(* IEC 61131-3 sources: plc-st-coding-agent/agent_dev/tests/samples, 4 files *)

(* ---- _bad_missing_clip.st ---- *)
FUNCTION_BLOCK FB
VAR_INPUT
    enable : BOOL;
    values : ARRAY[1..8] OF INT;
    count : INT;
    avgEnable : BOOL;
END_VAR
VAR_OUTPUT
    avgOut : REAL;
END_VAR
VAR
    i : INT;
    sum : DINT;
END_VAR
IF enable AND avgEnable AND count > 0 THEN
    sum := 0;
    FOR i := 1 TO count DO
        sum := sum + values[i];
    END_FOR
    avgOut := DINT_TO_REAL(sum) / INT_TO_REAL(count);
END_IF
END_FUNCTION_BLOCK

(* ---- bad_counter.st ---- *)
FUNCTION_BLOCK Bad
VAR_INPUT
    Start : BOOL;
END_VAR
VAR_OUTPUT
    Count : INT;
END_VAR
VAR
    Edge : BOOL;
END_VAR

IF Start THEN
    Count := Count + 1;
    Start := FALSE;
END_IF
IF Count > 100 THEN
    Edge := TRUE
END_IF;
IF Edge THEN
    Count := lalala + 1;
END_IF;
END_FUNCTION_BLOCK

(* ---- ok_counter.st ---- *)
FUNCTION_BLOCK Counter
VAR_INPUT
    Start : BOOL;
    Reset : BOOL;
END_VAR
VAR_OUTPUT
    Count : INT;
    Running : BOOL;
END_VAR
VAR
    prev : BOOL := FALSE;
END_VAR

IF Reset THEN
    Count := 0;
    Running := FALSE;
ELSIF Start AND NOT prev THEN
    Count := Count + 1;
    Running := TRUE;
END_IF;
prev := Start;
END_FUNCTION_BLOCK

(* ---- self_easy_01_ref.st ---- *)
FUNCTION_BLOCK FB
VAR_INPUT
    enable : BOOL;
    values : ARRAY[1..8] OF INT;
    count : INT;
    avgEnable : BOOL;
END_VAR
VAR_OUTPUT
    avgOut : REAL;
END_VAR
VAR
    i : INT;
    n : INT;
    sum : DINT;
END_VAR

(* 缓存语义见 Interpreter：输出变量在两次扫描之间保持上一次的值，
   enable / avgEnable / count=0 分支不写 avgOut，就自然"保持上一周期"。 *)

(* 先把有效样本数裁剪到 [0, 8]：count 为负或超过数组长度都不能越界 *)
n := count;
IF n < 0 THEN
    n := 0;
ELSIF n > 8 THEN
    n := 8;
END_IF

(* n = 0 时整段跳过，避免除零；avgOut 保持上一周期的值 *)
IF enable AND avgEnable AND n > 0 THEN
    sum := 0;
    FOR i := 1 TO n DO
        sum := sum + values[i];
    END_FOR
    avgOut := DINT_TO_REAL(sum) / INT_TO_REAL(n);
END_IF
END_FUNCTION_BLOCK
